SUBAPPLICATION Uebung_267_AX (* FIFO mit Adapter: Tastendruecke puffern, Q1 blinkt je Wert einmal (PROCESSED-Handshake) *)
  (* Standard: 61499-2; Description: Copyright (c) 2026 Meisterschulen am Ostbahnhof This program and the accompanying materials are made available under the terms of the Eclipse Public License 2.0 which is available at https://www.eclipse.org/legal/epl-2.0/ SPDX-License-Identifier: EPL-2.0 *)
  (* Version 1.0, 2026-11-08, Franz Höpfinger, Meisterschulen am Ostbahnhof, initial API and implementation and/or initial documentation *)
  PACKAGE Uebungen;
  IMPORT logiBUS::io::DI::logiBUS_DI::Input_I1;
  IMPORT logiBUS::io::DI::logiBUS_DI::Input_I4;
  IMPORT logiBUS::io::DI::logiBUS_DI_Events::BUTTON_SINGLE_CLICK;
  IMPORT logiBUS::io::DQ::logiBUS_DO::Output_Q1;
  IMPORT logiBUS::io::DQ::logiBUS_DO::Output_Q2;
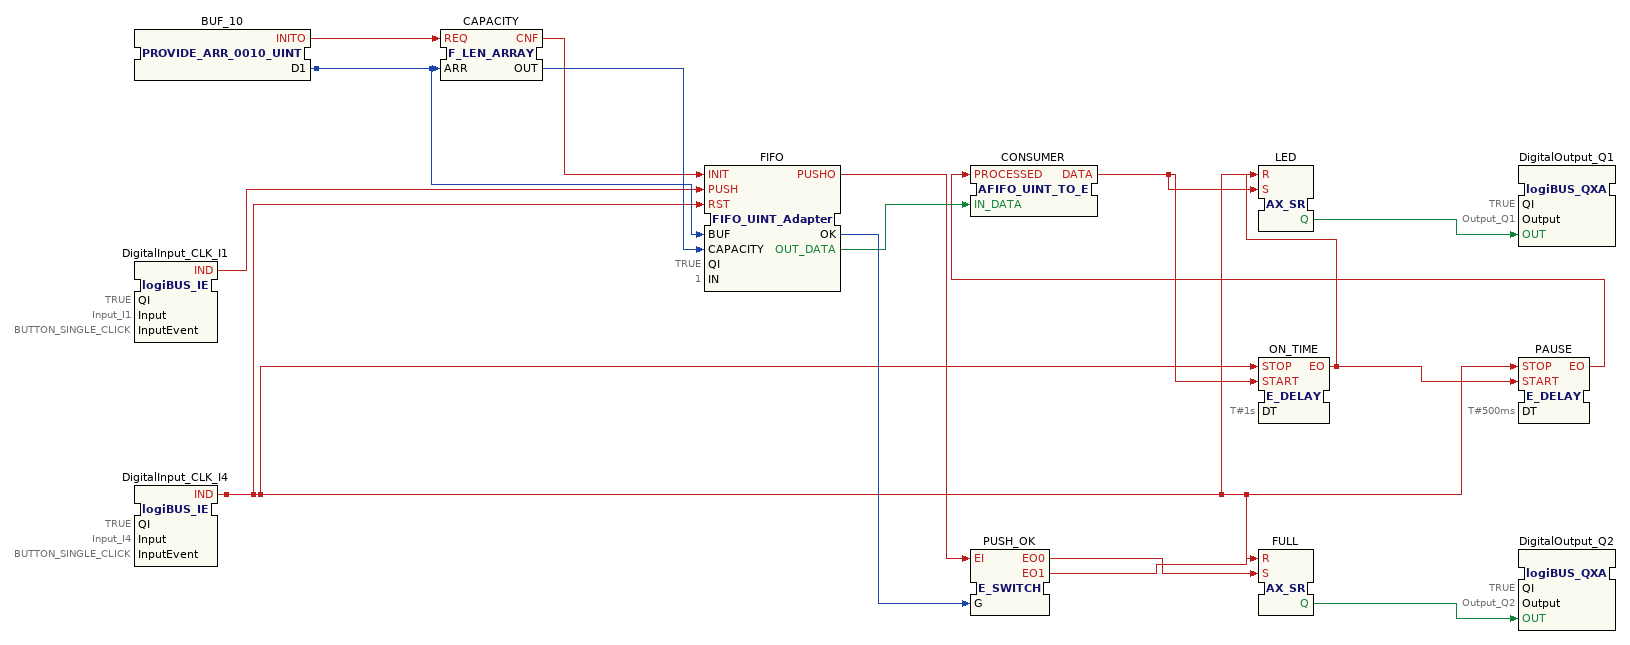
  FBS
    BUF_10 : eclipse4diac::convert::providers::PROVIDE_ARR_0010_UINT;
    CAPACITY : eclipse4diac::utils::arrays::F_LEN_ARRAY;
    FIFO : FIFO_adapter::FIFO_UINT_Adapter(QI := TRUE, IN := 1);
    CONSUMER : FIFO_adapter::AFIFO_UINT_TO_E;
    DigitalInput_CLK_I1 : logiBUS::io::DI::logiBUS_IE(QI := TRUE, Input := Input_I1, InputEvent := BUTTON_SINGLE_CLICK);
    DigitalInput_CLK_I4 : logiBUS::io::DI::logiBUS_IE(QI := TRUE, Input := Input_I4, InputEvent := BUTTON_SINGLE_CLICK);
    LED : adapter::events::unidirectional::AX_SR;
    ON_TIME : iec61499::events::E_DELAY(DT := T#1s);
    PAUSE : iec61499::events::E_DELAY(DT := T#500ms);
    DigitalOutput_Q1 : logiBUS::io::DQ::logiBUS_QXA(QI := TRUE, Output := Output_Q1);
    PUSH_OK : iec61499::events::E_SWITCH;
    FULL : adapter::events::unidirectional::AX_SR;
    DigitalOutput_Q2 : logiBUS::io::DQ::logiBUS_QXA(QI := TRUE, Output := Output_Q2);
  END_FBS
  EVENT_CONNECTIONS
    BUF_10.INITO TO CAPACITY.REQ;
    CAPACITY.CNF TO FIFO.INIT;
    DigitalInput_CLK_I1.IND TO FIFO.PUSH;
    DigitalInput_CLK_I4.IND TO FIFO.RST;
    DigitalInput_CLK_I4.IND TO ON_TIME.STOP;
    DigitalInput_CLK_I4.IND TO PAUSE.STOP;
    DigitalInput_CLK_I4.IND TO LED.R;
    DigitalInput_CLK_I4.IND TO FULL.R;
    CONSUMER.DATA TO LED.S;
    CONSUMER.DATA TO ON_TIME.START;
    ON_TIME.EO TO LED.R;
    ON_TIME.EO TO PAUSE.START;
    PAUSE.EO TO CONSUMER.PROCESSED;
    FIFO.PUSHO TO PUSH_OK.EI;
    PUSH_OK.EO0 TO FULL.S;
    PUSH_OK.EO1 TO FULL.R;
  END_CONNECTIONS
  DATA_CONNECTIONS
    BUF_10.D1 TO CAPACITY.ARR;
    BUF_10.D1 TO FIFO.BUF;
    CAPACITY.OUT TO FIFO.CAPACITY;
    FIFO.OK TO PUSH_OK.G;
  END_CONNECTIONS
  ADAPTER_CONNECTIONS
    FIFO.OUT_DATA TO CONSUMER.IN_DATA;
    LED.Q TO DigitalOutput_Q1.OUT;
    FULL.Q TO DigitalOutput_Q2.OUT;
  END_CONNECTIONS
END_SUBAPPLICATION
